(* PLC project g_conveyor_interlock_clean, Anonymous Benchmark Suite 1.0 *)
(* stored: creationDateTime 2026-07-09T00:00:00 *)

PROGRAM g_conveyor_interlock_clean
  VAR_INPUT
    run_cmd : BOOL;
    estop : BOOL;
    guard_open : BOOL;
    maint : BOOL;
  END_VAR
  VAR_OUTPUT
    conveyor : BOOL;
    warn : BOOL;
  END_VAR

(* LD diagram, written out as Structured Text *)
conveyor := NOT estop AND run_cmd AND NOT guard_open;
warn := estop;
END_PROGRAM

CONFIGURATION Config0
  RESOURCE Res0 ON PLC
    TASK tcyclic(INTERVAL := T#10ms, PRIORITY := 0);
    PROGRAM inst0 WITH tcyclic : g_conveyor_interlock_clean;
  END_RESOURCE
END_CONFIGURATION
